(* PLC project cycle, ESBMC probe 1.0 *)
(* stored: creationDateTime 2026-10-07T00:00:00 *)

PROGRAM cycle
  VAR_INPUT
    a : BOOL;
    b : BOOL;
    c : BOOL;
  END_VAR
  VAR_OUTPUT
    y : BOOL;
  END_VAR

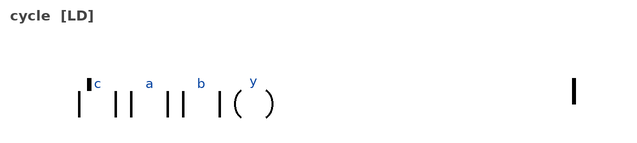
(* LD diagram, written out as Structured Text *)
y := (c OR FALSE (*loop*)) AND a AND b;
END_PROGRAM

CONFIGURATION Config0
  RESOURCE Res0 ON PLC
    TASK tcyclic(INTERVAL := T#10ms, PRIORITY := 0);
    PROGRAM inst0 WITH tcyclic : cycle;
  END_RESOURCE
END_CONFIGURATION
